TYPE "DT_PAR_GEN_SPEED"
VERSION : 0.1
   STRUCT
      STANDSTILL { S7_SetPoint := 'False'} : "DT_PARAM_SOLO" := (FALSE, 352, 0, 10.0, 0, T#0MS, 0.0, 0.0, '%');
      BRAKE { S7_SetPoint := 'False'} : "DT_PARAM_SOLO" := (FALSE, 353, 0, 15.0, 0, T#0MS, 0.0, 0.0, '%');
      EXCITATION { S7_SetPoint := 'False'} : "DT_PARAM_SOLO" := (FALSE, 354, 0, 95.0, 0, T#0MS, 0.0, 0.0, '%');
      SYNC { S7_SetPoint := 'False'} : "DT_PARAM_SOLO" := (FALSE, 355, 0, 98.0, 0, T#0MS, 0.0, 0.0, '%');
      OVERSPEED_1 { S7_SetPoint := 'False'} : "DT_PARAM_SOLO" := (FALSE, 356, 0, 110.0, 0, T#0MS, 0.0, 0.0, '%');
      OVERSPEED_2 { S7_SetPoint := 'False'} : "DT_PARAM_SOLO" := (FALSE, 357, 0, 120.0, 0, T#0MS, 0.0, 0.0, '%');
      STANDSTILL_HYST { S7_SetPoint := 'False'} : "DT_PARAM_SOLO" := (FALSE, 358, 0, 2.0, 0, T#0MS, 0.0, 0.0, '%');
      BRAKE_HYST { S7_SetPoint := 'False'} : "DT_PARAM_SOLO" := (FALSE, 359, 0, 2.0, 0, T#0MS, 0.0, 0.0, '%');
      EXCITATION_HYST { S7_SetPoint := 'False'} : "DT_PARAM_SOLO" := (FALSE, 360, 0, 5.0, 0, T#0MS, 0.0, 0.0, '%');
      SYNC_HYST { S7_SetPoint := 'False'} : "DT_PARAM_SOLO" := (FALSE, 361, 0, 5.0, 0, T#0MS, 0.0, 0.0, '%');
      OVERSPEED_1_HYST { S7_SetPoint := 'False'} : "DT_PARAM_SOLO" := (FALSE, 362, 0, 5.0, 0, T#0MS, 0.0, 0.0, '%');
      OVERSPEED_2_HYST { S7_SetPoint := 'False'} : "DT_PARAM_SOLO" := (FALSE, 363, 0, 5.0, 0, T#0MS, 0.0, 0.0, '%');
      PARAM_108 { S7_SetPoint := 'False'} : "DT_PARAM_SOLO" := (FALSE, 364, 0, 0.0, 0, T#0MS, 0.0, 0.0, '');
      PARAM_109 { S7_SetPoint := 'False'} : "DT_PARAM_SOLO" := (FALSE, 365, 0, 0.0, 0, T#0MS, 0.0, 0.0, '');
      PARAM_110 { S7_SetPoint := 'False'} : "DT_PARAM_SOLO" := (FALSE, 366, 0, 0.0, 0, T#0MS, 0.0, 0.0, '');
      PARAM_111 { S7_SetPoint := 'False'} : "DT_PARAM_SOLO" := (FALSE, 367, 0, 0.0, 0, T#0MS, 0.0, 0.0, '');
      MAIN_SPEED_VAL_LOW { S7_SetPoint := 'False'} : "DT_PARAM_SOLO" := (FALSE, 368, 0, 0.0, 0, T#0MS, 0.0, 0.0, 'rpm');
      MAIN_SPEED_VAL_HIGH { S7_SetPoint := 'False'} : "DT_PARAM_SOLO" := (FALSE, 369, 0, 1500.0, 0, T#0MS, 0.0, 0.0, 'rpm');
      MAIN_SPEED_SCAL_FACTOR { S7_SetPoint := 'False'} : "DT_PARAM_SOLO" := (FALSE, 370, 0, 1.0, 0, T#0MS, 0.0, 0.0, '-');
      MAIN_SPEED_OFFSET { S7_SetPoint := 'False'} : "DT_PARAM_SOLO" := (FALSE, 371, 0, 0.0, 0, T#0MS, 0.0, 0.0, 'rpm');
      RED_SPEED_VAL_LOW { S7_SetPoint := 'False'} : "DT_PARAM_SOLO" := (FALSE, 372, 0, 0.0, 0, T#0MS, 0.0, 0.0, 'rpm');
      RED_SPEED_VAL_HIGH { S7_SetPoint := 'False'} : "DT_PARAM_SOLO" := (FALSE, 373, 0, 1500.0, 0, T#0MS, 0.0, 0.0, 'rpm');
      RED_SPEED_SCAL_FACTOR { S7_SetPoint := 'False'} : "DT_PARAM_SOLO" := (FALSE, 374, 0, 1.0, 0, T#0MS, 0.0, 0.0, '-');
      RED_SPEED_OFFSET { S7_SetPoint := 'False'} : "DT_PARAM_SOLO" := (FALSE, 375, 0, 0.0, 0, T#0MS, 0.0, 0.0, 'rpm');
      PARAM_120 { S7_SetPoint := 'False'} : "DT_PARAM_SOLO" := (FALSE, 376, 0, 0.0, 0, T#0MS, 0.0, 0.0, '');
      PARAM_121 { S7_SetPoint := 'False'} : "DT_PARAM_SOLO" := (FALSE, 377, 0, 0.0, 0, T#0MS, 0.0, 0.0, '');
      PARAM_122 { S7_SetPoint := 'False'} : "DT_PARAM_SOLO" := (FALSE, 378, 0, 0.0, 0, T#0MS, 0.0, 0.0, '');
      PARAM_123 { S7_SetPoint := 'False'} : "DT_PARAM_SOLO" := (FALSE, 379, 0, 0.0, 0, T#0MS, 0.0, 0.0, '');
      PARAM_124 { S7_SetPoint := 'False'} : "DT_PARAM_SOLO" := (FALSE, 380, 0, 0.0, 0, T#0MS, 0.0, 0.0, '');
      PARAM_125 { S7_SetPoint := 'False'} : "DT_PARAM_SOLO" := (FALSE, 381, 0, 0.0, 0, T#0MS, 0.0, 0.0, '');
      PARAM_126 { S7_SetPoint := 'False'} : "DT_PARAM_SOLO" := (FALSE, 382, 0, 0.0, 0, T#0MS, 0.0, 0.0, '');
      PARAM_127 { S7_SetPoint := 'False'} : "DT_PARAM_SOLO" := (FALSE, 383, 0, 0.0, 0, T#0MS, 0.0, 0.0, '');
   END_STRUCT;

END_TYPE

